FUNCTION_BLOCK Draining
VAR_INPUT
	diEnabled : BOOL;
END_VAR
VAR_OUTPUT
	doEnabled : BOOL;
END_VAR
VAR_IN_OUT
	DrainingPhase : TPhaseDraining;
	DrainingValve : TValve;
END_VAR
VAR
END_VAR

{region "Aut/Man"}
    // switching state of engine - automatic or manual control (default state is manual)
  	IF DrainingPhase.Cmd.ManCtrl THEN
      	DrainingPhase.State.ManCtrl := TRUE;
		DrainingPhase.State.AutCtrl := FALSE;
	ELSIF DrainingPhase.Cmd.AutCtrl THEN
        DrainingPhase.State.ManCtrl := FALSE;
		DrainingPhase.State.AutCtrl := TRUE; 
    END_IF;
		 
	IF (NOT DrainingPhase.State.AutCtrl AND NOT DrainingPhase.State.ManCtrl) THEN
		DrainingPhase.State.ManCtrl := TRUE;
	END_IF

	DrainingPhase.Cmd.ManCtrl := FALSE;
	DrainingPhase.Cmd.AutCtrl := FALSE;
{endregion}

{region "ManCtrl"}
    // processing manual actions - if command is processed, it is sets to FALSE even if can't be processed
    // Phase commands are start, stop, pause and resume 
    // Start - open draining valve 
    // Stop - close draining valve
    // Pause - close draining valve
    // Resume - open draining valve
    // real states of phase are writed into states in phase structure
    IF DrainingPhase.State.ManCtrl THEN
		IF DrainingPhase.State.Idle AND DrainingPhase.Cmd.StartMan THEN
			DrainingPhase.State.Running := TRUE;
			DrainingPhase.State.Idle := FALSE;
			DrainingPhase.State.Paused := FALSE;
		 	DrainingPhase.State.Done := FALSE;
		ELSIF DrainingPhase.Cmd.StopMan THEN
			DrainingPhase.State.Running := FALSE;
			DrainingPhase.State.Idle := TRUE;
			DrainingPhase.State.Paused := FALSE;
		ELSIF DrainingPhase.State.Running AND DrainingPhase.Cmd.PauseMan THEN
			DrainingPhase.State.Running := FALSE;
			DrainingPhase.State.Idle := FALSE;
			DrainingPhase.State.Paused := TRUE;
		ELSIF DrainingPhase.State.Paused AND DrainingPhase.Cmd.ResumeMan THEN
			DrainingPhase.State.Running := TRUE;
			DrainingPhase.State.Idle := FALSE;
			DrainingPhase.State.Paused := FALSE;
			DrainingPhase.State.Done := FALSE;
		END_IF
    END_IF;
	
	DrainingPhase.Cmd.StartMan := FALSE;
	DrainingPhase.Cmd.StopMan := FALSE;
	DrainingPhase.Cmd.PauseMan := FALSE;
	DrainingPhase.Cmd.ResumeMan := FALSE;
{endregion}

{region "AutCtrl"}
    //if request to run in automatic mode -> set auto request to open of filling valve to 1 and close to 0, if not open 0 close 1
    // commands should be sets to false after their processing
    IF DrainingPhase.State.AutCtrl THEN
		IF DrainingPhase.State.Idle AND DrainingPhase.Cmd.StartAut THEN
			DrainingPhase.State.Running := TRUE;
			DrainingPhase.State.Idle := FALSE;
		 	DrainingPhase.State.Done := FALSE;
		ELSIF DrainingPhase.Cmd.StopAut THEN
			DrainingPhase.State.Running := FALSE;
			DrainingPhase.State.Idle := TRUE;
			DrainingPhase.State.Paused := FALSE;
		END_IF
    END_IF;
	
	DrainingPhase.Cmd.StartAut := FALSE;
	DrainingPhase.Cmd.StopAut := FALSE;
{endregion}
{region "Done"}
    //every phase should have finish condition - draining phase - if water level is below requested level
    //after that done state should be setted to 1
    IF DrainingPhase.State.Running AND (DrainingPhase.WaterLevel <= DrainingPhase.ParamDrainLevel) THEN // edit based on speed of simulation 
        DrainingPhase.Cmd.StopMan := TRUE;
        DrainingPhase.Cmd.StopAut := TRUE;
        DrainingPhase.State.Done := TRUE;
    END_IF;

    IF DrainingPhase.Cmd.ResetDone THEN
        DrainingPhase.State.Done := FALSE;
        DrainingPhase.Cmd.ResetDone := FALSE;
    END_IF;
{endregion}

{region "States"} 
    //Command valve in cases of states
    IF DrainingPhase.State.Running THEN
        DrainingValve.Cmd.Req2OpenAut := TRUE;
        DrainingValve.Cmd.Req2CloseAut := FALSE;
    ELSE
        DrainingValve.Cmd.Req2OpenAut := FALSE;
        DrainingValve.Cmd.Req2CloseAut := TRUE;
    END_IF;
{endregion}

// delault state of phase - if not any state sets state to idle
IF (NOT DrainingPhase.State.Idle) AND (NOT DrainingPhase.State.Paused) AND (NOT DrainingPhase.State.Running) THEN
    DrainingPhase.State.Idle := 1;
END_IF;

// write binary states into int value for visualization
IF DrainingPhase.State.Idle THEN
    DrainingPhase.State.StateInt := Global.PhIdle;
ELSIF DrainingPhase.State.Running THEN
    DrainingPhase.State.StateInt := Global.PhRunning;
ELSE
    DrainingPhase.State.StateInt := Global.PhPause;
END_IF;

//Ponechte pro moznost retezeni volani bloku v LAD
doEnabled := diEnabled;

END_FUNCTION_BLOCK

(* stored: Version 1.1.0.1, ProductVersion 3.1.4026.21
   POU Draining: Id {a501d01f-bc41-415b-8bb8-19a7a35d7bf8}, SpecialFunc None *)
